// TIA Portal V20 export
DATA_BLOCK "T5_Datos"   // DB42900
{ S7_Optimized_Access := 'TRUE' }
AUTHOR : IA
FAMILY : PRUEBA
VERSION : 0.1
// Tanda 1b: datos
// stored: AutoNumber false
   VAR
      Tog : Bool;   // Cambia cada ciclo
      Falso : Bool := false;
      Int_0 : Int := 0;
      Int_1 : Int := 1;
      Int_3 : Int := 3;
      Int_4 : Int := 4;
      Int_5 : Int := 5;
      Int_9 : Int := 9;
      Int_10 : Int := 10;
      Int_20 : Int := 20;
      Int_50 : Int := 50;
      Int_100 : Int := 100;
      Real_2 : Real := 2.0;
      Real_0_5 : Real := 0.5;
      Real_16 : Real := 16.0;
      UInt_2 : UInt := 2;
      UInt_3 : UInt := 3;
      DWord_00F0 : DWord := 16#000000F0;
      Arr_A : Array[0..9] of Int;
      Arr_B : Array[0..9] of Int;
      Arr_C : Array[0..9] of Int;
      Arr_E : Array[0..9] of Int;
      Inc_Var : Int;
      Dec_Var : Int;
      MIN_Out : Int;
      MAX_Out : Int;
      LIMIT_Out : Int;
      Expt_Out : Real;
      DECO_Out : DWord;
      ENCO_Out : Int;
      SEL_Out : Int;
      OK_Q : Bool;
      NOK_Q : Bool;
      R_TRIG_Q : Bool;
      F_TRIG_Q : Bool;
      RS_Mem : Bool;
      RS_Q : Bool;
      Bits_BF : Array[0..7] of Bool;
      Bits_RBF : Array[0..7] of Bool;
      Arr_F : Array[0..9] of Int;
      Arr_U : Array[0..9] of Int;
      UInt_10 : UInt := 10;
      MBV_Ret : Int;
      UDInt_2 : UDInt := 2;
      DInt_0 : DInt := 0;
      DInt_5 : DInt := 5;
      NORM_Out : Real;
      SCALE_Out : Int;
   END_VAR
BEGIN
END_DATA_BLOCK
